// Mitsubishi GX Works2 project: Test2   PLC: Q06UDEH

PROGRAM MAIN
VAR
  HPR : POINTER;
  H_HPR : POINTER;
END_VAR
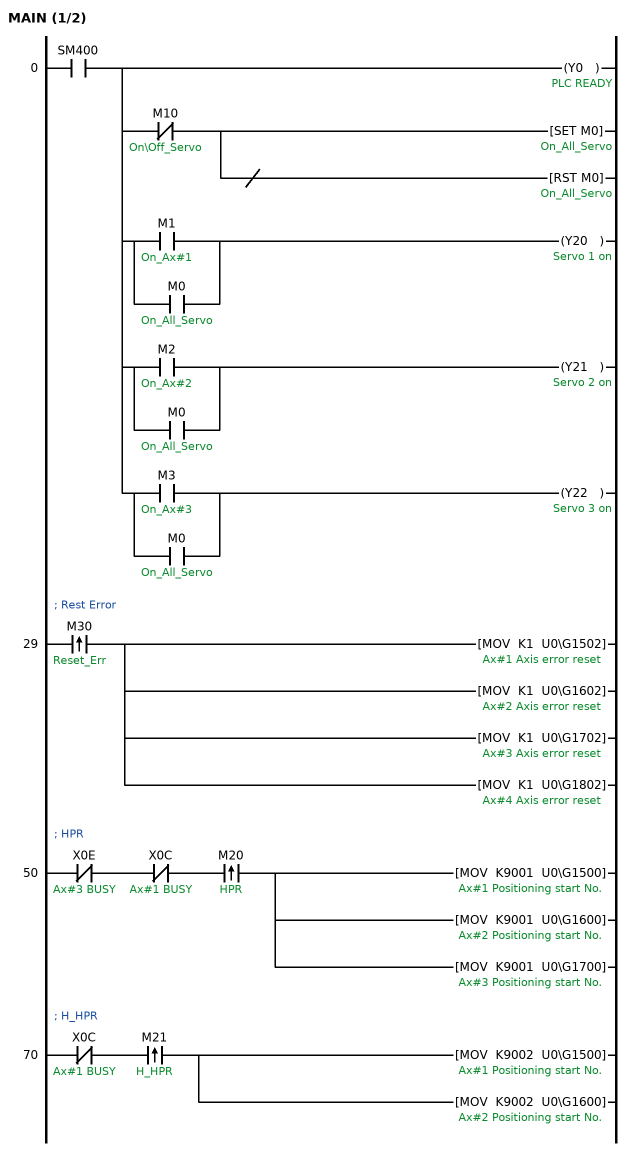
0     LD      SM400
      OUT     Y0  ; PLC READY
      MPS
      ANI     M10  ; On\Off_Servo
      SET     M0  ; On_All_Servo
      INV
      RST     M0  ; On_All_Servo
      MRD
      LD      M1  ; On_Ax#1
      OR      M0  ; On_All_Servo
      ANB
      OUT     Y20  ; Servo 1 on
      MRD
      LD      M2  ; On_Ax#2
      OR      M0  ; On_All_Servo
      ANB
      OUT     Y21  ; Servo 2 on
      MPP
      LD      M3  ; On_Ax#3
      OR      M0  ; On_All_Servo
      ANB
      OUT     Y22  ; Servo 3 on
; Rest Error
29    LDP     M30  ; Reset_Err
      MOV     K1 U0\G1502  ; Ax#1 Axis error reset
      MOV     K1 U0\G1602  ; Ax#2 Axis error reset
      MOV     K1 U0\G1702  ; Ax#3 Axis error reset
      MOV     K1 U0\G1802  ; Ax#4 Axis error reset
; HPR
50    LDI     X0E  ; Ax#3 BUSY
      ANI     X0C  ; Ax#1 BUSY
      ANDP    M20  ; HPR
      MOV     K9001 U0\G1500  ; Ax#1 Positioning start No.
      MOV     K9001 U0\G1600  ; Ax#2 Positioning start No.
      MOV     K9001 U0\G1700  ; Ax#3 Positioning start No.
; H_HPR
70    LDI     X0C  ; Ax#1 BUSY
      ANDP    M21  ; H_HPR
      MOV     K9002 U0\G1500
      MOV     K9002 U0\G1600
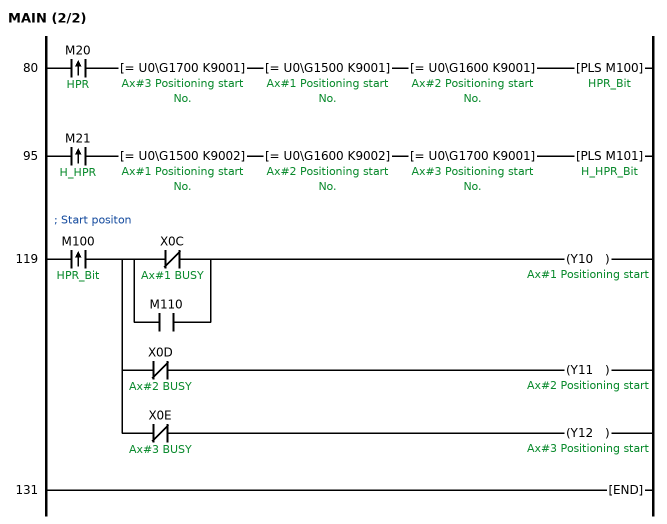
80    LDP     M20  ; HPR
      AND=    U0\G1700 K9001  ; Ax#3 Positioning start No.
      AND=    U0\G1500 K9001  ; Ax#1 Positioning start No.
      AND=    U0\G1600 K9001  ; Ax#2 Positioning start No.
      PLS     M100  ; HPR_Bit
95    LDP     M21  ; H_HPR
      AND=    U0\G1500 K9002  ; Ax#1 Positioning start No.
      AND=    U0\G1600 K9002  ; Ax#2 Positioning start No.
      AND=    U0\G1700 K9001  ; Ax#3 Positioning start No.
      PLS     M101  ; H_HPR_Bit
; Start positon
119   LDP     M100  ; HPR_Bit
      MPS
      LDI     X0C  ; Ax#1 BUSY
      OR      M110
      ANB
      OUT     Y10  ; Ax#1 Positioning start
      MRD
      ANI     X0D  ; Ax#2 BUSY
      OUT     Y11  ; Ax#2 Positioning start
      MPP
      ANI     X0E  ; Ax#3 BUSY
      OUT     Y12  ; Ax#3 Positioning start
131   END
END_PROGRAM

PROGRAM Tracking
VAR
  bInit : BOOL;  (* Cờ khởi tạo chu trình ban đầu *)
  bM100_Old : BOOL;  (* Lưu trạng thái M100 để bắt cạnh lên *)
  bMCode_Handled : BOOL;  (* Cờ chống kích trùng van keo tại Point 2 *)
  bQd75Ready : BOOL;  (* Giám sát trạng thái module QD75 *)
  iState : INT;  (* Máy trạng thái FSM (0, 10, 20, 30, 40, 50) *)
  dErrCode : INT;  (* Mã lỗi chẩn đoán phần mềm *)
  wAxis1_Err : INT;  (* Đọc mã lỗi phần cứng Trục 1 (Md.23) *)
  wAxis2_Err : INT;  (* Đọc mã lỗi phần cứng Trục 2 (Md.23) *)
  wAxis3_Err : INT;  (* Đọc mã lỗi phần cứng Trục 3 (Md.23) *)
  dTarget_X_Sync : DINT;  (* Tọa độ kết thúc trượt Trục X ($Target_X + \Delta X$) *)
  Target_X : DINT;  (* Tọa độ đón đầu đỉnh Trục X ($0.1\ \mu\text{m}$) *)
  Target_Y : DINT;  (* Tọa độ đỉnh Trục Y ($0.1\ \mu\text{m}$) *)
  Target_Z_Down : DINT;  (* Độ cao hạ kim để xả keo ($0.1\ \mu\text{m}$) *)
  Speed_Approach : DINT;  (* Vận tốc bay nội suy tiếp cận ($0.01\text{ mm/min}$) *)
  Speed_Sync : DINT;  (* Vận tốc đồng tốc trục X khi xả keo *)
  DeltaX_Sync : DINT;  (* Quãng đường trượt đồng tốc ($0.1\ \mu\text{m}$) *)
  Target_Z_Safe : DINT;  (* Độ cao an toàn rút kim ($0.0\text{ mm} = 0$) *)
  Vertex_Index : INT;  (* Số thứ tự đỉnh (1..4) *)
  Cmd_Start_Vertex : BOOL;  (* Lệnh kích chạy đỉnh từ TwinCAT 3 *)
  Ack_Vertex_Done : BOOL;  (* Báo hoàn thành đỉnh về TwinCAT 3 *)
  Robot_Busy : BOOL;  (* Cờ báo Gantry đang chuyển động *)
  Robot_In_Position : BOOL;  (* Cờ báo Gantry đã vào đích *)
  Robot_Alarm : BOOL;  (* Cờ báo động lỗi hệ thống *)
  Cmd_Cycle_Reset : BOOL;  (* Lệnh dừng khẩn cấp / Hủy chu trình *)
  Valve_Internal : BOOL;  (* Cuộn nội bộ điều khiển van keo *)
  Valve_Output : BOOL;  (* Ngõ ra Transistor vật lý mở van keo (Slot 1) *)
  bReq_Start_Y10 : BOOL;
  bValve_Timer_Run : BOOL;
END_VAR
(***************************************************************************************************)
(* PROGRAM: Tracking (ST) - BẢN FIX 0 CẢNH BÁO, 0 DOUBLE-COIL                                      *)
(***************************************************************************************************)

(* 1. KHỞI TẠO NỘI BỘ *)
IF SM402 OR NOT bInit THEN
    iState := 0;
    dErrCode := 0;
    dTarget_X_Sync := 0;
    bReq_Start_Y10 := FALSE;
    bMCode_Handled := FALSE;
    bInit := TRUE;
END_IF;

bQd75Ready := X0;

(* 2. DỪNG KHẨN CẤP / RESET *)
IF Cmd_Cycle_Reset THEN
    iState := 0;
    bReq_Start_Y10 := FALSE;
    bMCode_Handled := FALSE;
END_IF;

(* 3. ĐỌC MÃ LỖI MODULE QD75 *)
FROM(TRUE, H0, 806, 1, wAxis1_Err);
FROM(TRUE, H0, 906, 1, wAxis2_Err);
FROM(TRUE, H0, 1006, 1, wAxis3_Err);

IF Cmd_Cycle_Reset AND (X8 OR X9 OR XA) THEN
    TO(TRUE, 1, H0, 1502, 1);
    TO(TRUE, 1, H0, 1602, 1);
    TO(TRUE, 1, H0, 1702, 1);
    dErrCode := 0;
END_IF;

(* 4. MÁY TRẠNG THÁI FSM *)
CASE iState OF

    0: (* IDLE *)
        bReq_Start_Y10 := FALSE;
        IF Cmd_Start_Vertex AND NOT bM100_Old THEN
            IF X0 AND NOT XC AND NOT XD AND NOT XE AND NOT X8 AND NOT X9 AND NOT XA AND NOT Cmd_Cycle_Reset THEN
                iState := 10;
                dErrCode := 0;
            ELSE
                dErrCode := 901;
            END_IF;
        END_IF;

    10: (* PRE-CHECK & NẠP BUFFER *)
        dTarget_X_Sync := Target_X + DeltaX_Sync;
        
        IF (Target_X < 0) OR (Target_X > 1800000) OR (dTarget_X_Sync < 0) OR (dTarget_X_Sync > 1800000) THEN
            dErrCode := 501;
            iState := 0;
        ELSIF (Target_Y < 0) OR (Target_Y > 1700000) THEN
            dErrCode := 502;
            iState := 0;
        ELSIF (Target_Z_Down < 0) OR (Target_Z_Down > 520000) OR (Target_Z_Safe < 0) OR (Target_Z_Safe > 520000) OR (Target_Z_Down < Target_Z_Safe) THEN
            dErrCode := 503;
            iState := 0;
        ELSE
            (* POINT 1 *)
            TO(TRUE, 16#1503, H0, 2000, 1);
            TO(TRUE, 0, H0, 2001, 1);
            DTO(TRUE, 0, H0, 2002, 1);
            DTO(TRUE, Speed_Approach, H0, 2004, 1);
            DTO(TRUE, Target_X, H0, 2006, 1);
            DTO(TRUE, Target_Y, H0, 8006, 1);
            DTO(TRUE, Target_Z_Down, H0, 14006, 1);

            (* POINT 2 *)
            TO(TRUE, 16#1503, H0, 2010, 1);
            TO(TRUE, 1, H0, 2011, 1);
            DTO(TRUE, 0, H0, 2012, 1);
            DTO(TRUE, Speed_Sync, H0, 2014, 1);
            DTO(TRUE, dTarget_X_Sync, H0, 2016, 1);
            DTO(TRUE, Target_Y, H0, 8016, 1);
            DTO(TRUE, Target_Z_Down, H0, 14016, 1);

            (* POINT 3 *)
            TO(TRUE, 16#1500, H0, 2020, 1);
            TO(TRUE, 0, H0, 2021, 1);
            DTO(TRUE, 0, H0, 2022, 1);
            DTO(TRUE, Speed_Approach, H0, 2024, 1);
            DTO(TRUE, dTarget_X_Sync, H0, 2026, 1);
            DTO(TRUE, Target_Y, H0, 8026, 1);
            DTO(TRUE, Target_Z_Safe, H0, 14026, 1);

            TO(TRUE, 1, H0, 1500, 1); (* Cd.3 = 1 *)
            iState := 20;
        END_IF;

    20: (* YÊU CẦU START *)
        bReq_Start_Y10 := TRUE;
        IF X10 THEN
            bReq_Start_Y10 := FALSE;
            iState := 30;
        END_IF;

    30: (* CHẠY & BƠM KEO *)
        IF X4 AND NOT bMCode_Handled THEN
            bMCode_Handled := TRUE;
            TO(TRUE, 1, H0, 1504, 1); (* Cd.7 = 1 xóa cờ X4 *)
        END_IF;
        
        IF NOT X4 THEN
            TO(TRUE, 0, H0, 1504, 1);
        END_IF;
        
        IF X14 AND NOT XC AND NOT XD AND NOT XE THEN
            bMCode_Handled := FALSE;
            iState := 40;
        END_IF;

    40: (* HOÀN THÀNH ĐỈNH *)
        iState := 50;

    50: (* CHỜ MASTER HẠ M100 *)
        IF NOT Cmd_Start_Vertex THEN
            iState := 0;
        END_IF;

END_CASE;

(* 5. ĐỊNH THÌ VAN KEO 30MS TỐC ĐỘ CAO *)
bValve_Timer_Run := (iState = 30) AND bMCode_Handled AND NOT TS0;
TIMER_H_M(bValve_Timer_Run, TC0, 3);

(***************************************************************************************************)
(* 6. TẦNG XUẤT COIL DUY NHẤT (MỖI COIL CHỈ XUẤT ĐÚNG 1 LẦN -> TRIỆT TIÊU 100% CẢNH BÁO)            *)
(***************************************************************************************************)
Robot_Busy := (iState >= 10) AND (iState <= 30) AND NOT Cmd_Cycle_Reset;
Robot_In_Position := (iState = 40) OR (iState = 50);
Ack_Vertex_Done := (iState = 40) OR (iState = 50);
Robot_Alarm := X8 OR X9 OR XA OR (dErrCode <> 0);

(* Lệnh dừng trục hãm khẩn: gán duy nhất 1 lần *)
Y4 := Cmd_Cycle_Reset;
Y5 := Cmd_Cycle_Reset;
Y6 := Cmd_Cycle_Reset;

(* Lệnh Start Trục 1: Xuất ra bit trung gian M110 để không đè cuộn Y10 của MAIN *)
M110 := bReq_Start_Y10 AND NOT Cmd_Cycle_Reset;

(* Van keo vật lý Y20: gán duy nhất 1 lần *)
Valve_Output := bValve_Timer_Run AND NOT Cmd_Cycle_Reset;

bM100_Old := Cmd_Start_Vertex;
END_PROGRAM

// device comments not shown above
X0  ; QD75 READY
X4  ; Ax#1 M code ON
X8  ; Ax#1 Error detection
X9  ; Ax#2 Error detection
X0A  ; Ax#3 Error detection
X10  ; Ax#1 Start complete
X14  ; Ax#1 Positioning complete
Y4  ; Axis #1 Axis stop
Y5  ; Axis #2 Axis stop
Y6  ; Axis #3 Axis stop
X1  ; Synchronization flag signal
X5  ; Ax#2 M code ON
X6  ; Ax#3 M code ON
X7  ; Ax#4 M code ON
X0B  ; Ax#4 Error detection
X0F  ; Ax#4 BUSY
X11  ; Ax#2 Start complete
X12  ; Ax#3 Start complete
X13  ; Ax#4 Start complete
X15  ; Ax#2 Positioning complete
X16  ; Ax#3 Positioning complete
X17  ; Ax#4 Positioning complete
Y7  ; Axis #4 Axis stop
Y8  ; Ax#1 Forward run JOG start
Y9  ; Ax#1 Reverse run JOG start
Y0A  ; Ax#2 Forward run JOG start
Y0B  ; Ax#2 Reverse run JOG start
Y0C  ; Ax#3 Forward run JOG start
Y0D  ; Ax#3 Reverse run JOG start
Y0E  ; Ax#4 Forward run JOG start
Y0F  ; Ax#4 Reverse run JOG start
Y13  ; Ax#4 Positioning start
Y14  ; Ax#1 Exe prhbtn flag sgnl
Y15  ; Ax#2 Exe prhbtn flag sgnl
Y16  ; Ax#3 Exe prhbtn flag sgnl
Y17  ; Ax#4 Exe prhbtn flag sgnl
Y23  ; Open Brk
M1000  ; Trigger 1 phoi
M2000  ; Lenh diem keo
M3000  ; Báo FIFO đầy
D1200  ; Tọa độ X bám thực tế gửi sang Ro
D2200  ; Tọa độ Y bám thực tế gửi sang Ro
R0  ; X tam camera mm
R2  ; Y tam camera mm
R4  ; Goc xoay 0.1 do
R6  ; Toc bang mm/s live
R8  ; Z bay 0.1mm giu
R10  ; Z cham 0.1mm giu
R12  ; Toc chay
R14  ; Toc do max
